Fanuc KAREL source: KA00065.KL

PROGRAM KA00065
%NOLOCKGROUP
VAR
  SRC: XYZWPR
  DST: POSITION
BEGIN
  SRC.X = 1.0
  DST = SRC
END KA00065
